FUNCTION_BLOCK CipSequence_AOI (* Migrated from IEC 61131-3 ST *)
  (* Standard: 61499-2 *)
  (* Version 1.0, 2026-11-06, st2fb *)
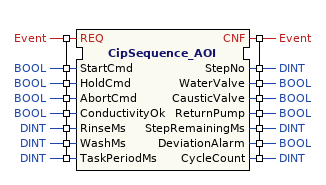
  EVENT_INPUT
    REQ WITH StartCmd, HoldCmd, AbortCmd, ConductivityOk, RinseMs, WashMs, TaskPeriodMs;
  END_EVENT
  EVENT_OUTPUT
    CNF WITH StepNo, WaterValve, CausticValve, ReturnPump, StepRemainingMs, DeviationAlarm, CycleCount;
  END_EVENT
  VAR_INPUT
    StartCmd : BOOL;
    HoldCmd : BOOL;
    AbortCmd : BOOL;
    ConductivityOk : BOOL;
    RinseMs : DINT;
    WashMs : DINT;
    TaskPeriodMs : DINT;
  END_VAR
  VAR_OUTPUT
    StepNo : DINT;
    WaterValve : BOOL;
    CausticValve : BOOL;
    ReturnPump : BOOL;
    StepRemainingMs : DINT;
    DeviationAlarm : BOOL;
    CycleCount : DINT;
  END_VAR
  VAR
    StepTimer_EN : BOOL := FALSE;
    StepTimer_TT : BOOL := FALSE;
    StepTimer_DN : BOOL := FALSE;
    StepTimer_ACC : DINT := 0;
    StepTimer_PRE : DINT := 0;
    StepTimer_ENABLE : BOOL := FALSE;
    DevTimer_EN : BOOL := FALSE;
    DevTimer_TT : BOOL := FALSE;
    DevTimer_DN : BOOL := FALSE;
    DevTimer_ACC : DINT := 0;
    DevTimer_PRE : DINT := 0;
    DevTimer_ENABLE : BOOL := FALSE;
    OS_PREV : BOOL := FALSE;
    OS_OUT : BOOL := FALSE;
    Preset : DINT := 0;
  END_VAR
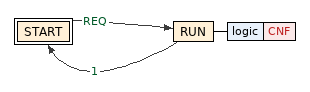
  EC_STATES
    START;
    RUN : logic -> CNF;
  END_STATES
  EC_TRANSITIONS
    START TO RUN := REQ;
    RUN TO START := 1;
  END_TRANSITIONS
  ALGORITHM logic IN ST:
OS_OUT := StartCmd AND NOT OS_PREV;
OS_PREV := StartCmd;

WaterValve := FALSE;
CausticValve := FALSE;
ReturnPump := FALSE;

IF AbortCmd THEN
  StepNo := 0;
  StepTimer_ACC := 0;
  StepTimer_EN := FALSE;
  StepTimer_TT := FALSE;
  StepTimer_DN := FALSE;
END_IF;

CASE StepNo OF
  0:
    Preset := RinseMs;
    IF OS_OUT AND NOT AbortCmd THEN
      StepNo := 10;
    END_IF;
  10:
    WaterValve := TRUE;
    ReturnPump := TRUE;
    IF StepTimer_DN THEN
      StepTimer_ACC := 0;
      StepTimer_EN := FALSE;
      StepTimer_TT := FALSE;
      StepTimer_DN := FALSE;
      Preset := WashMs;
      StepNo := 20;
    END_IF;
  20:
    CausticValve := TRUE;
    ReturnPump := TRUE;
    IF StepTimer_DN THEN
      StepTimer_ACC := 0;
      StepTimer_EN := FALSE;
      StepTimer_TT := FALSE;
      StepTimer_DN := FALSE;
      Preset := RinseMs;
      StepNo := 30;
    END_IF;
  30:
    WaterValve := TRUE;
    ReturnPump := TRUE;
    IF StepTimer_DN THEN
      StepTimer_ACC := 0;
      StepTimer_EN := FALSE;
      StepTimer_TT := FALSE;
      StepTimer_DN := FALSE;
      CycleCount := CycleCount + 1;
      StepNo := 0;
    END_IF;
END_CASE;

StepTimer_ENABLE := (StepNo = 10 OR StepNo = 30 OR (StepNo = 20 AND ConductivityOk)) AND NOT HoldCmd;
StepTimer_PRE := Preset;
IF StepTimer_ENABLE AND StepTimer_EN AND NOT StepTimer_DN THEN
  StepTimer_ACC := StepTimer_ACC + TaskPeriodMs;
  IF StepTimer_ACC >= StepTimer_PRE THEN
    StepTimer_ACC := StepTimer_PRE;
    StepTimer_DN := TRUE;
  END_IF;
END_IF;
IF NOT StepTimer_ENABLE THEN
  StepTimer_ACC := 0;
  StepTimer_DN := FALSE;
END_IF;
StepTimer_EN := StepTimer_ENABLE;
StepTimer_TT := StepTimer_EN AND NOT StepTimer_DN;
StepRemainingMs := Preset - StepTimer_ACC;

DevTimer_ENABLE := (StepNo = 20) AND NOT ConductivityOk;
DevTimer_PRE := 200;
IF DevTimer_ENABLE AND DevTimer_EN AND NOT DevTimer_DN THEN
  DevTimer_ACC := DevTimer_ACC + TaskPeriodMs;
  IF DevTimer_ACC >= DevTimer_PRE THEN
    DevTimer_ACC := DevTimer_PRE;
    DevTimer_DN := TRUE;
  END_IF;
END_IF;
IF NOT DevTimer_ENABLE THEN
  DevTimer_ACC := 0;
  DevTimer_DN := FALSE;
END_IF;
DevTimer_EN := DevTimer_ENABLE;
DevTimer_TT := DevTimer_EN AND NOT DevTimer_DN;
DeviationAlarm := DevTimer_DN;
  END_ALGORITHM
END_FUNCTION_BLOCK
